(* IEC 61131-3 sources: sis-interlock-demo/tests/POUs/TruthTables/FB_VoteTableRig, 9 files *)

(* ---- FB_VoteTableRig.decl.st ---- *)
// AUTO-GENERATED by tools_project/gen_voting_tests.py — не редактировать: правьте генератор или модель
//   tools_project/vote_model.py и запустите python tools_project/gen_voting_tests.py
// Назначение: стенд таблиц истинности голосования: строка таблицы → входы F_VoteEval или
//             FB_Voting → байт результата по разделу 12.2. Ожидаемые байты считает модель.
// Автор:      kr0nsch; код — генератор tools_project/gen_voting_tests.py
// Версия:     0.1.0
// Документ:   docs/DESIGN.md, раздел «12.2 Таблицы истинности (генерируются)»
// ВНИМАНИЕ:   код демонстрационный и не предназначен для систем безопасности. Реальная ПАЗ
//             требует определения SIL, сертифицированных аппаратных и программных средств
//             и валидации по ГОСТ Р МЭК 61511.
FUNCTION_BLOCK FB_VoteTableRig
VAR
    fbTime : PL.FB_FakeTime;    // время стоит (LTIME#1H): байпасы не истекают
    fbVote : FB_Voting;         // ФБ под тестом (уровень 2)
    stIn   : ST_VoteIn;         // входы строки
    stCmd  : ST_VoteCmd;        // запросы байпаса строки
    stCfg  : ST_VotingCfg;      // конфигурация таблицы (раздел 12.2)
END_VAR

(* ---- Encode.method.decl.st ---- *)
// AUTO-GENERATED by tools_project/gen_voting_tests.py — не редактировать: правьте генератор или модель
//   tools_project/vote_model.py и запустите python tools_project/gen_voting_tests.py
// Ожидаемый байт (раздел 12.2): бит 0 — xTrip, бит 1 — xDegraded, биты 2–4 — индекс eArchEff
// (0 — None, 1 — 1oo1, 2 — 1oo2, 3 — 2oo2, 4 — 2oo3, 5 — ForcedTrip, 7 — вне перечисления),
// биты 5–7 — действующие байпасы каналов 1..3
METHOD Encode : BYTE
VAR_INPUT
    xTrip     : BOOL;            // требование срабатывания
    xDegraded : BOOL;            // деградация
    eArchEff  : E_VoteArch;      // действующая схема
    bBypass   : BYTE;            // действующие байпасы: бит k-1 — канал k
END_VAR
VAR
    bCode : BYTE;                // результат
END_VAR

(* ---- Encode.method.impl.st ---- *)
// AUTO-GENERATED by tools_project/gen_voting_tests.py — не редактировать: правьте генератор или модель
//   tools_project/vote_model.py и запустите python tools_project/gen_voting_tests.py
CASE eArchEff OF
    E_VoteArch.None:
        bCode := 0;
    E_VoteArch.Vote1oo1:
        bCode := 1;
    E_VoteArch.Vote1oo2:
        bCode := 2;
    E_VoteArch.Vote2oo2:
        bCode := 3;
    E_VoteArch.Vote2oo3:
        bCode := 4;
    E_VoteArch.ForcedTrip:
        bCode := 5;
ELSE
    bCode := 7;
END_CASE
bCode := SHL(bCode, 2) OR SHL(bBypass, 5);
IF xTrip THEN
    bCode := bCode OR 16#01;
END_IF
IF xDegraded THEN
    bCode := bCode OR 16#02;
END_IF
Encode := bCode;

(* ---- EvalRow.method.decl.st ---- *)
// AUTO-GENERATED by tools_project/gen_voting_tests.py — не редактировать: правьте генератор или модель
//   tools_project/vote_model.py и запустите python tools_project/gen_voting_tests.py
// Строка уровня 1: состояние канала k — код (uiRow SHR 2(k-1)) AND 3: 0 — Normal, 1 — Demand,
// 2 — Invalid, 3 — Bypassed; каналы k > N — NotUsed. Результат — байт Encode
METHOD EvalRow : BYTE
VAR_INPUT
    uiRow : UINT;                // номер строки
END_VAR
VAR
    aeCh  : ARRAY[1..GVL_Const.SIS_VOTE_CH_MAX] OF E_ChannelState;   // состояния каналов строки
    wRow  : WORD;                // номер строки как битовая строка
    wCode : WORD;                // код состояния канала
    uiK   : UINT;                // номер канала
    uiN   : UINT;                // каналов в схеме
    stRes : ST_VoteResult;       // результат F_VoteEval
END_VAR

(* ---- EvalRow.method.impl.st ---- *)
// AUTO-GENERATED by tools_project/gen_voting_tests.py — не редактировать: правьте генератор или модель
//   tools_project/vote_model.py и запустите python tools_project/gen_voting_tests.py
uiN := F_VoteArchChannels(eArch := stCfg.eArch);
wRow := UINT_TO_WORD(uiRow);
FOR uiK := 1 TO GVL_Const.SIS_VOTE_CH_MAX DO
    IF uiK <= uiN THEN
        wCode := SHR(wRow, 2 * (uiK - 1)) AND 16#0003;
        CASE WORD_TO_UINT(wCode) OF
            0:
                aeCh[uiK] := E_ChannelState.Normal;
            1:
                aeCh[uiK] := E_ChannelState.Demand;
            2:
                aeCh[uiK] := E_ChannelState.Invalid;
        ELSE
            aeCh[uiK] := E_ChannelState.Bypassed;
        END_CASE
    ELSE
        aeCh[uiK] := E_ChannelState.NotUsed;
    END_IF
END_FOR
stRes := F_VoteEval(eArch := stCfg.eArch, ePolicy := stCfg.ePolicy, aeCh := aeCh);
EvalRow := Encode(xTrip := stRes.xTrip, xDegraded := stRes.xDegraded, eArchEff := stRes.eArchEff, bBypass := 0);

(* ---- FbRow.method.decl.st ---- *)
// AUTO-GENERATED by tools_project/gen_voting_tests.py — не редактировать: правьте генератор или модель
//   tools_project/vote_model.py и запустите python tools_project/gen_voting_tests.py
// Строка уровня 2: для канала k биты b = 3(k-1): b — требование (DI: axDi := FALSE; AI: 60.0,
// иначе 40.0), b+1 — достоверность, b+2 — запрос байпаса. Два вызова одного экземпляра: со снятыми
// запросами байпаса (сбрасывает байпасы прошлой строки) и с полной строкой. Результат — байт Encode
METHOD FbRow : BYTE
VAR_INPUT
    uiRow : UINT;                // номер строки
END_VAR
VAR
    wRow    : WORD;              // номер строки как битовая строка
    uiK     : UINT;              // номер канала
    uiN     : UINT;              // каналов в схеме
    uiShift : UINT;              // номер бита требования канала
    xDem    : BOOL;              // требование канала
    xValid  : BOOL;              // достоверность канала
    axReq   : ARRAY[1..GVL_Const.SIS_VOTE_CH_MAX] OF BOOL;   // запросы байпаса строки
    bBypass : BYTE;              // действующие байпасы: бит k-1 — канал k
END_VAR

(* ---- FbRow.method.impl.st ---- *)
// AUTO-GENERATED by tools_project/gen_voting_tests.py — не редактировать: правьте генератор или модель
//   tools_project/vote_model.py и запустите python tools_project/gen_voting_tests.py
uiN := F_VoteArchChannels(eArch := stCfg.eArch);
wRow := UINT_TO_WORD(uiRow);
FOR uiK := 1 TO GVL_Const.SIS_VOTE_CH_MAX DO
    uiShift := 3 * (uiK - 1);
    xDem := (uiK <= uiN) AND ((SHR(wRow, uiShift) AND 16#0001) <> 0);
    xValid := (uiK <= uiN) AND ((SHR(wRow, uiShift + 1) AND 16#0001) <> 0);
    axReq[uiK] := (uiK <= uiN) AND ((SHR(wRow, uiShift + 2) AND 16#0001) <> 0);
    stIn.axDi[uiK] := NOT xDem;
    stIn.axDiValid[uiK] := xValid;
    IF xDem THEN
        stIn.arAi_eu[uiK] := 60.0;
    ELSE
        stIn.arAi_eu[uiK] := 40.0;
    END_IF
    stIn.axAiValid[uiK] := xValid;
    stCmd.axBypassReq[uiK] := FALSE;
END_FOR
fbVote(stIn := stIn, stCmd := stCmd, stCfg := stCfg, xBypassPermit := TRUE, uiCause := 1, itfTime := fbTime);
FOR uiK := 1 TO GVL_Const.SIS_VOTE_CH_MAX DO
    stCmd.axBypassReq[uiK] := axReq[uiK];
END_FOR
fbVote(stIn := stIn, stCmd := stCmd, stCfg := stCfg, xBypassPermit := TRUE, uiCause := 1, itfTime := fbTime);
bBypass := 0;
FOR uiK := 1 TO GVL_Const.SIS_VOTE_CH_MAX DO
    IF fbVote.stSts.aeBypass[uiK] = E_BypassState.Active THEN
        bBypass := bBypass OR SHL(BYTE#1, uiK - 1);
    END_IF
END_FOR
FbRow := Encode(xTrip := fbVote.xTrip, xDegraded := fbVote.stSts.xDegraded, eArchEff := fbVote.stSts.eArchEff,
    bBypass := bBypass);

(* ---- Setup.method.decl.st ---- *)
// AUTO-GENERATED by tools_project/gen_voting_tests.py — не редактировать: правьте генератор или модель
//   tools_project/vote_model.py и запустите python tools_project/gen_voting_tests.py
// Конфигурация таблицы по разделу 12.2: уставка 50.0 (High), гистерезис и рассогласование
// выключены, tBypassMax = T#1H, uiMaxBypass = MIN(1, N - 1), xDiHealthy = TRUE
METHOD Setup
VAR_INPUT
    eArch   : E_VoteArch;        // схема
    ePolicy : E_DegradePolicy;   // политика
    eInput  : E_SisInputKind;    // вид входов (для уровня 1 не действует)
END_VAR

(* ---- Setup.method.impl.st ---- *)
// AUTO-GENERATED by tools_project/gen_voting_tests.py — не редактировать: правьте генератор или модель
//   tools_project/vote_model.py и запустите python tools_project/gen_voting_tests.py
stCfg.eArch := eArch;
stCfg.ePolicy := ePolicy;
stCfg.eInput := eInput;
stCfg.xDiHealthy := TRUE;
stCfg.eLimitDir := E_LimitDir.High;
stCfg.rTripLimit_eu := 50.0;
stCfg.rHyst_eu := 0.0;
stCfg.rDiscrepancyMax_eu := 0.0;
stCfg.tDiscrepancyDelay := T#0S;
stCfg.tBypassMax := T#1H;
IF F_VoteArchChannels(eArch := eArch) > 1 THEN
    stCfg.uiMaxBypass := 1;
ELSE
    stCfg.uiMaxBypass := 0;
END_IF
